// TIA Portal V20 export
// export: Created 2026-10-19T18:03:08.52848Z, ExportSetting WithDefaults, DisplayName Totally Integrated Automation Portal, DisplayVersion V20 Update 6, DisplayName TIA Portal Openness, DisplayVersion V20 Update 6, DisplayName TIA Portal Version Control Interface, DisplayVersion V20 Update 6, DisplayName SINAMICS Startdrive Advanced, DisplayVersion V20 SP1, DisplayName SINAMICS Startdrive G130, G150, S120, S150, SINAMICS MV, G220, S200, S210, DisplayVersion V20 SP1, DisplayName SINAMICS Startdrive G110M, G120, G120C, G120D, G120P, G115D, DisplayVersion V20 SP1, DisplayName STEP 7 Professional, DisplayVersion V20 Update 6, DisplayName STEP 7 Safety, DisplayVersion V20 Update 2, DisplayName WinCC Basic/Comfort/Advanced, DisplayVersion V20 Update 6, DisplayName WinCC Unified, DisplayVersion V20 Update 6
DATA_BLOCK "SB_Alarm"   // DB118
{ S7_Optimized_Access := 'TRUE' }
VERSION : 0.1
// stored: AutoNumber true, DBAccessibleFromOPCUA true, DBAccessibleFromWebserver true, InstanceOfName SAI_SB_Alarm, InstanceOfType UDT, IsOnlyStoredInLoadMemory false, IsWriteProtectedInAS false
"SAI_SB_Alarm"
   // VAR
   //    "LC overload in operation range" : Bool;
   //    "LC Mix" : Bool;
   //    "Application defined 1" : Bool;
   //    "Application defined 2" : Bool;
   //    "Application defined 3" : Bool;
   //    "Application defined 4" : Bool;
   //    "Application defined 5" : Bool;
   //    "Application defined 7" : Bool;
   //    "Rate of change error" : Bool;
   //    "Communication error" : Bool;
   //    "Over / under voltage" : Bool;
   //    "Weight drift" : Bool;
   //    Breach : Bool;
   //    "Calibration expired" : Bool;
   //    "Over Current" : Bool;
   //    "LC overload in normal range" : Bool;
   // END_VAR
BEGIN
END_DATA_BLOCK
